// TIA Portal V20 export
// export: Created 2026-10-19T18:45:31.9794258Z, ExportSetting None, DisplayName Totally Integrated Automation Portal, DisplayVersion V20 Update 6, DisplayName TIA Portal Openness, DisplayVersion V20 Update 6, DisplayName TIA Portal Version Control Interface, DisplayVersion V20 Update 6, DisplayName SINAMICS Startdrive Advanced, DisplayVersion V20 SP1, DisplayName SINAMICS Startdrive G130, G150, S120, S150, SINAMICS MV, G220, S200, S210, DisplayVersion V20 SP1, DisplayName SINAMICS Startdrive G110M, G120, G120C, G120D, G120P, G115D, DisplayVersion V20 SP1, DisplayName STEP 7 Professional, DisplayVersion V20 Update 6, DisplayName STEP 7 Safety, DisplayVersion V20 Update 2, DisplayName WinCC Basic/Comfort/Advanced, DisplayVersion V20 Update 6, DisplayName WinCC Unified, DisplayVersion V20 Update 6
VAR_GLOBAL   // PLC tag table "IO_Turck_2"
   "Light_Bar_2_Percent_Width1(2)" AT %QB657 : Byte;   // Last byte - 16
   "Light_Bar_2_Bounce_Style(2)" AT %QB659 : Byte;   // Last byte - 14
   "Light_Bar_1_Color1(2)" AT %QB633 : Byte;   // Last byte - 2
   "Light_Bar_1_Intensity2(2)" AT %QB623 : Byte;   // Last byte - 12
   "Light_Bar_1_Color2(2)" AT %QB625 : Byte;   // Last byte - 10
   "Light_Bar_1_Animation(2)" AT %QB635 : Byte;   // Last byte
   "Light_Bar_2_Color2(2)" AT %QB663 : Byte;   // Last byte - 10
   "Light_Bar_2_Animation(2)" AT %QB673 : Byte;   // Last byte
   "Light_Bar_2_Direction(2)" AT %QB655 : Byte;   // Last byte - 18
   "Light_Bar_1_Intensity1(2)" AT %QB631 : Byte;   // Last byte - 4
   "Light_Bar_2_Intensity1(2)" AT %QB669 : Byte;   // Last byte - 4
   "Light_Bar_2_Color1(2)" AT %QB671 : Byte;   // Last byte - 2
   "Light_Bar_2_Pulse_Pattern(2)" AT %QB665 : Byte;   // Last byte - 8
   "Light_Bar_2_Speed(2)" AT %QB667 : Byte;   // Last byte - 6
   "Light_Bar_1_Pulse_Pattern(2)" AT %QB627 : Byte;   // Last byte - 8
   "Light_Bar_2_Intensity2(2)" AT %QB661 : Byte;   // Last byte - 12
   "Light_Bar_1_Percent_Width1(2)" AT %QB619 : Byte;   // Last byte - 16
   "Light_Bar_1_Speed(2)" AT %QB629 : Byte;   // Last byte - 6
   "Light_Bar_1_Bounce_Style(2)" AT %QB621 : Byte;   // Last byte - 14
   "Light_Bar_1_1_Direction(2)" AT %QB617 : Byte;   // Last byte - 18
END_VAR
